Fanuc KAREL source: kx00028.compact.KL

PROGRAM KX00028
%STACKSIZE=65535
%PRIORITY=65535
%TIMESLICE=8
%NOLOCKGROUP
VAR
I : INTEGER
J : INTEGER
B : BOOLEAN
F : FILE
S : STRING[80]
P : XYZWPR
BEGIN
I=1
END KX00028
